// TIA Portal V19 export
TYPE "ST_PLACE_POSITION"
   STRUCT
      Place : Array[0..50] of "ST_Pos";
   END_STRUCT;
END_TYPE
